Staubli VAL3: appLauncher.dtx

bool _bAtHome
bool _bEndCycle
bool _bHeavyAlarm
bool _bIsScara
bool _bShowEndBt
bool _bShowPauseBt
bool _bShowResetBt
bool _bShowStartBt
bool _bShowStopBt
bool bBool
bool bControlByRobot = true
bool bTosave
frame test3 = {fatherId=world[0]}
num _nAvgCapacity
num _nBestCapacity
num _nCTIndex
num _nCapacity
num _nClock[10]
  [1] = 12488.271809
  [3] = 12488.271821
num _nCycleTime[10]
num _nLastStateCMD
num _nOmacStat
num _nStateCMD
num nCycleCmd
num nErrorCode = 1
num nLastLib
num nProgCode
string _sArmType
string _sOmacCmd
string _sOmacStatus = "1"
string _sPageAvergeCapacity
string _sPageBestCapacity
string _sPageCurrentCapacity
string _sPageCycleStatus
string _sPageHerej
string _sPagePosition
string _sPageProfile
string _sPageRobotStatus
string _sPageSN
string sMsg
num nForce[6]
public bool bGetMovId
mdesc mHome = {accel=20, vel=20, decel=20, blend=off}
string sSessionList
pointRx pPowerOFF = {fatherId=world[0]}
bool bMemState
pointRx pHere1 = {fatherId=world[0]}
pointRx pHere2 = {fatherId=world[0]}
bool bAutoConnectMove
